(* PLC project Vn_ton_call_edit_pt, Beckhoff Automation GmbH TwinCAT PLC Control 3.5.13.21 *)
(* stored: creationDateTime 1970-01-01T00:00:00 *)

PROGRAM Vn_ton_call_edit_pt

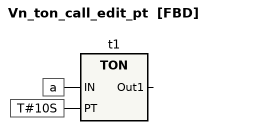
(* FBD diagram, written out as Structured Text *)
t1(IN := a, PT := T#10S);
END_PROGRAM
